       IF #inB15 THEN
           #outR15 := #inR15 * 2.0;
       END_IF;
       // step 536
       #tI36 := #inI16 + #cI26;
       IF #inB16 THEN
           #outR16 := #inR16 * 2.0;
       END_IF;
       // step 537
       #tI37 := #inI17 + #cI27;
       IF #inB17 THEN
           #outR17 := #inR17 * 2.0;
       END_IF;
       // step 538
       #tI38 := #inI18 + #cI28;
       IF #inB18 THEN
           #outR18 := #inR18 * 2.0;
       END_IF;
       // step 539
       #tI39 := #inI19 + #cI29;
       IF #inB19 THEN
           #outR19 := #inR19 * 2.0;
       END_IF;
       // step 540
       #tI40 := #inI20 + #cI0;
       IF #inB20 THEN
           #outR0 := #inR0 * 2.0;
       END_IF;
       // step 541
       #tI41 := #inI21 + #cI1;
       IF #inB21 THEN
           #outR1 := #inR1 * 2.0;
       END_IF;
       // step 542
       #tI42 := #inI22 + #cI2;
       IF #inB22 THEN
           #outR2 := #inR2 * 2.0;
       END_IF;
       // step 543
       #tI43 := #inI23 + #cI3;
       IF #inB23 THEN
           #outR3 := #inR3 * 2.0;
       END_IF;
       // step 544
       #tI44 := #inI24 + #cI4;
       IF #inB24 THEN
           #outR4 := #inR4 * 2.0;
       END_IF;
       // step 545
       #tI45 := #inI25 + #cI5;
       IF #inB25 THEN
           #outR5 := #inR5 * 2.0;
       END_IF;
       // step 546
       #tI46 := #inI26 + #cI6;
       IF #inB26 THEN
           #outR6 := #inR6 * 2.0;
       END_IF;
       // step 547
       #tI47 := #inI27 + #cI7;
       IF #inB27 THEN
           #outR7 := #inR7 * 2.0;
       END_IF;
       // step 548
       #tI48 := #inI28 + #cI8;
       IF #inB28 THEN
           #outR8 := #inR8 * 2.0;
       END_IF;
       // step 549
       #tI49 := #inI29 + #cI9;
       IF #inB29 THEN
           #outR9 := #inR9 * 2.0;
       END_IF;
       END_REGION
       REGION part 11
       // step 550
       #tI50 := #inI30 + #cI10;
       IF #inB30 THEN
           #outR10 := #inR10 * 2.0;
       END_IF;
       // step 551
       #tI51 := #inI31 + #cI11;
       IF #inB31 THEN
           #outR11 := #inR11 * 2.0;
       END_IF;
       // step 552
       #tI52 := #inI32 + #cI12;
       IF #inB32 THEN
           #outR12 := #inR12 * 2.0;
       END_IF;
       // step 553
       #tI53 := #inI33 + #cI13;
       IF #inB33 THEN
           #outR13 := #inR13 * 2.0;
       END_IF;
       // step 554
       #tI54 := #inI34 + #cI14;
       IF #inB34 THEN
           #outR14 := #inR14 * 2.0;
       END_IF;
       // step 555
       #tI55 := #inI35 + #cI15;
       IF #inB35 THEN
           #outR15 := #inR15 * 2.0;
       END_IF;
       // step 556
       #tI56 := #inI36 + #cI16;
       IF #inB36 THEN
           #outR16 := #inR16 * 2.0;
       END_IF;
       // step 557
       #tI57 := #inI37 + #cI17;
       IF #inB37 THEN
           #outR17 := #inR17 * 2.0;
       END_IF;
       // step 558
       #tI58 := #inI38 + #cI18;
       IF #inB38 THEN
           #outR18 := #inR18 * 2.0;
       END_IF;
       // step 559
       #tI59 := #inI39 + #cI19;
       IF #inB39 THEN
           #outR19 := #inR19 * 2.0;
       END_IF;
       // step 560
       #tI60 := #inI0 + #cI20;
       IF #inB0 THEN
           #outR0 := #inR0 * 2.0;
       END_IF;
       // step 561
       #tI61 := #inI1 + #cI21;
       IF #inB1 THEN
           #outR1 := #inR1 * 2.0;
       END_IF;
       // step 562
       #tI62 := #inI2 + #cI22;
       IF #inB2 THEN
           #outR2 := #inR2 * 2.0;
       END_IF;
       // step 563
       #tI63 := #inI3 + #cI23;
       IF #inB3 THEN
           #outR3 := #inR3 * 2.0;
       END_IF;
       // step 564
       #tI64 := #inI4 + #cI24;
       IF #inB4 THEN
           #outR4 := #inR4 * 2.0;
       END_IF;
       // step 565
       #tI65 := #inI5 + #cI25;
       IF #inB5 THEN
           #outR5 := #inR5 * 2.0;
       END_IF;
       // step 566
       #tI66 := #inI6 + #cI26;
       IF #inB6 THEN
           #outR6 := #inR6 * 2.0;
       END_IF;
       // step 567
       #tI67 := #inI7 + #cI27;
       IF #inB7 THEN
           #outR7 := #inR7 * 2.0;
       END_IF;
       // step 568
       #tI68 := #inI8 + #cI28;
       IF #inB8 THEN
           #outR8 := #inR8 * 2.0;
       END_IF;
       // step 569
       #tI69 := #inI9 + #cI29;
       IF #inB9 THEN
           #outR9 := #inR9 * 2.0;
       END_IF;
       // step 570
       #tI70 := #inI10 + #cI0;
       IF #inB10 THEN
           #outR10 := #inR10 * 2.0;
       END_IF;
       // step 571
       #tI71 := #inI11 + #cI1;
       IF #inB11 THEN
           #outR11 := #inR11 * 2.0;
       END_IF;
       // step 572
       #tI72 := #inI12 + #cI2;
       IF #inB12 THEN
           #outR12 := #inR12 * 2.0;
       END_IF;
       // step 573
       #tI73 := #inI13 + #cI3;
       IF #inB13 THEN
           #outR13 := #inR13 * 2.0;
       END_IF;
       // step 574
       #tI74 := #inI14 + #cI4;
       IF #inB14 THEN
           #outR14 := #inR14 * 2.0;
       END_IF;
       // step 575
       #tI75 := #inI15 + #cI5;
       IF #inB15 THEN
           #outR15 := #inR15 * 2.0;
       END_IF;
       // step 576
       #tI76 := #inI16 + #cI6;
       IF #inB16 THEN
           #outR16 := #inR16 * 2.0;
       END_IF;
       // step 577
       #tI77 := #inI17 + #cI7;
       IF #inB17 THEN
           #outR17 := #inR17 * 2.0;
       END_IF;
       // step 578
       #tI78 := #inI18 + #cI8;
       IF #inB18 THEN
           #outR18 := #inR18 * 2.0;
       END_IF;
       // step 579
       #tI79 := #inI19 + #cI9;
       IF #inB19 THEN
           #outR19 := #inR19 * 2.0;
       END_IF;
       // step 580
       #tI80 := #inI20 + #cI10;
       IF #inB20 THEN
           #outR0 := #inR0 * 2.0;
       END_IF;
       // step 581
       #tI81 := #inI21 + #cI11;
       IF #inB21 THEN
           #outR1 := #inR1 * 2.0;
       END_IF;
       // step 582
       #tI82 := #inI22 + #cI12;
       IF #inB22 THEN
           #outR2 := #inR2 * 2.0;
       END_IF;
       // step 583
       #tI83 := #inI23 + #cI13;
       IF #inB23 THEN
           #outR3 := #inR3 * 2.0;
       END_IF;
       // step 584
       #tI84 := #inI24 + #cI14;
       IF #inB24 THEN
           #outR4 := #inR4 * 2.0;
       END_IF;
       // step 585
       #tI85 := #inI25 + #cI15;
       IF #inB25 THEN
           #outR5 := #inR5 * 2.0;
       END_IF;
       // step 586
       #tI86 := #inI26 + #cI16;
       IF #inB26 THEN
           #outR6 := #inR6 * 2.0;
       END_IF;
       // step 587
       #tI87 := #inI27 + #cI17;
       IF #inB27 THEN
           #outR7 := #inR7 * 2.0;
       END_IF;
       // step 588
       #tI88 := #inI28 + #cI18;
       IF #inB28 THEN
           #outR8 := #inR8 * 2.0;
       END_IF;
       // step 589
       #tI89 := #inI29 + #cI19;
       IF #inB29 THEN
           #outR9 := #inR9 * 2.0;
       END_IF;
       // step 590
       #tI90 := #inI30 + #cI20;
       IF #inB30 THEN
           #outR10 := #inR10 * 2.0;
       END_IF;
       // step 591
       #tI91 := #inI31 + #cI21;
       IF #inB31 THEN
           #outR11 := #inR11 * 2.0;
       END_IF;
       // step 592
       #tI92 := #inI32 + #cI22;
       IF #inB32 THEN
           #outR12 := #inR12 * 2.0;
       END_IF;
       // step 593
       #tI93 := #inI33 + #cI23;
       IF #inB33 THEN
           #outR13 := #inR13 * 2.0;
       END_IF;
       // step 594
       #tI94 := #inI34 + #cI24;
       IF #inB34 THEN
           #outR14 := #inR14 * 2.0;
       END_IF;
       // step 595
       #tI95 := #inI35 + #cI25;
       IF #inB35 THEN
           #outR15 := #inR15 * 2.0;
       END_IF;
       // step 596
       #tI96 := #inI36 + #cI26;
       IF #inB36 THEN
           #outR16 := #inR16 * 2.0;
       END_IF;
       // step 597
       #tI97 := #inI37 + #cI27;
       IF #inB37 THEN
           #outR17 := #inR17 * 2.0;
       END_IF;
       // step 598
       #tI98 := #inI38 + #cI28;
       IF #inB38 THEN
           #outR18 := #inR18 * 2.0;
       END_IF;
       // step 599
       #tI99 := #inI39 + #cI29;
       IF #inB39 THEN
           #outR19 := #inR19 * 2.0;
       END_IF;
       END_REGION
END_FUNCTION_BLOCK

FUNCTION_BLOCK "FB_MixedStl"   // FB900, LAD
{ S7_Optimized_Access := 'TRUE' }
VERSION : 0.1
   VAR_INPUT
      inB0 : Bool;   // input bit 0
      inB1 : Bool;
      inB2 : Bool;
      inB3 : Bool;
      inB4 : Bool;
      inB5 : Bool;
      inB6 : Bool;
      inB7 : Bool;
      inB8 : Bool;
      inB9 : Bool;
      inB10 : Bool;   // input bit 10
      inB11 : Bool;
      inB12 : Bool;
      inB13 : Bool;
      inB14 : Bool;
      inB15 : Bool;
      inB16 : Bool;
      inB17 : Bool;
      inB18 : Bool;
      inB19 : Bool;
      inB20 : Bool;   // input bit 20
      inB21 : Bool;
      inB22 : Bool;
      inB23 : Bool;
      inB24 : Bool;
      inB25 : Bool;
      inB26 : Bool;
      inB27 : Bool;
      inB28 : Bool;
      inB29 : Bool;
      inB30 : Bool;   // input bit 30
      inB31 : Bool;
      inB32 : Bool;
      inB33 : Bool;
      inB34 : Bool;
      inB35 : Bool;
      inB36 : Bool;
      inB37 : Bool;
      inB38 : Bool;
      inB39 : Bool;
      inI0 : Int;
      inI1 : Int;
      inI2 : Int;
      inI3 : Int;
      inI4 : Int;
      inI5 : Int;
      inI6 : Int;
      inI7 : Int;
      inI8 : Int;
      inI9 : Int;
      inI10 : Int;
      inI11 : Int;
      inI12 : Int;
      inI13 : Int;
      inI14 : Int;
      inI15 : Int;
      inI16 : Int;
      inI17 : Int;
      inI18 : Int;
      inI19 : Int;
      inI20 : Int;
      inI21 : Int;
      inI22 : Int;
      inI23 : Int;
      inI24 : Int;
      inI25 : Int;
      inI26 : Int;
      inI27 : Int;
      inI28 : Int;
      inI29 : Int;
      inI30 : Int;
      inI31 : Int;
      inI32 : Int;
      inI33 : Int;
      inI34 : Int;
      inI35 : Int;
      inI36 : Int;
      inI37 : Int;
      inI38 : Int;
      inI39 : Int;
      inR0 : Real;
      inR1 : Real;
      inR2 : Real;
      inR3 : Real;
      inR4 : Real;
      inR5 : Real;
      inR6 : Real;
      inR7 : Real;
      inR8 : Real;
      inR9 : Real;
      inR10 : Real;
      inR11 : Real;
      inR12 : Real;
      inR13 : Real;
      inR14 : Real;
      inR15 : Real;
      inR16 : Real;
      inR17 : Real;
      inR18 : Real;
      inR19 : Real;
      inD0 : DInt;
      inD1 : DInt;
      inD2 : DInt;
      inD3 : DInt;
      inD4 : DInt;
      inD5 : DInt;
      inD6 : DInt;
      inD7 : DInt;
      inD8 : DInt;
      inD9 : DInt;
      inD10 : DInt;
      inD11 : DInt;
      inD12 : DInt;
      inD13 : DInt;
      inD14 : DInt;
      inD15 : DInt;
      inD16 : DInt;
      inD17 : DInt;
      inD18 : DInt;
      inD19 : DInt;
      inArr : Array[0..99] of Int;   // input array
      inStr : String[40];
      inSt : Struct
         x : Int;
         y : Real;
         z : Bool;
      END_STRUCT;
   END_VAR
   VAR_OUTPUT
      outB0 : Bool;
      outB1 : Bool;
      outB2 : Bool;
      outB3 : Bool;
      outB4 : Bool;
      outB5 : Bool;
      outB6 : Bool;
      outB7 : Bool;
      outB8 : Bool;
      outB9 : Bool;
      outB10 : Bool;
      outB11 : Bool;
      outB12 : Bool;
      outB13 : Bool;
      outB14 : Bool;
      outB15 : Bool;
      outB16 : Bool;
      outB17 : Bool;
      outB18 : Bool;
      outB19 : Bool;
      outB20 : Bool;
      outB21 : Bool;
      outB22 : Bool;
      outB23 : Bool;
      outB24 : Bool;
      outB25 : Bool;
      outB26 : Bool;
      outB27 : Bool;
      outB28 : Bool;
      outB29 : Bool;
      outB30 : Bool;
      outB31 : Bool;
      outB32 : Bool;
      outB33 : Bool;
      outB34 : Bool;
      outB35 : Bool;
      outB36 : Bool;
      outB37 : Bool;
      outB38 : Bool;
      outB39 : Bool;
      outI0 : Int;   // output int 0
      outI1 : Int;
      outI2 : Int;
      outI3 : Int;
      outI4 : Int;
      outI5 : Int;
      outI6 : Int;
      outI7 : Int;
      outI8 : Int;
      outI9 : Int;
      outI10 : Int;   // output int 10
      outI11 : Int;
      outI12 : Int;
      outI13 : Int;
      outI14 : Int;
      outI15 : Int;
      outI16 : Int;
      outI17 : Int;
      outI18 : Int;
      outI19 : Int;
      outI20 : Int;   // output int 20
      outI21 : Int;
      outI22 : Int;
      outI23 : Int;
      outI24 : Int;
      outI25 : Int;
      outI26 : Int;
      outI27 : Int;
      outI28 : Int;
      outI29 : Int;
      outI30 : Int;   // output int 30
      outI31 : Int;
      outI32 : Int;
      outI33 : Int;
      outI34 : Int;
      outI35 : Int;
      outI36 : Int;
      outI37 : Int;
      outI38 : Int;
      outI39 : Int;
      outR0 : Real;
      outR1 : Real;
      outR2 : Real;
      outR3 : Real;
      outR4 : Real;
      outR5 : Real;
      outR6 : Real;
      outR7 : Real;
      outR8 : Real;
      outR9 : Real;
      outR10 : Real;
      outR11 : Real;
      outR12 : Real;
      outR13 : Real;
      outR14 : Real;
      outR15 : Real;
      outR16 : Real;
      outR17 : Real;
      outR18 : Real;
      outR19 : Real;
      outD0 : DInt;
      outD1 : DInt;
      outD2 : DInt;
      outD3 : DInt;
      outD4 : DInt;
      outD5 : DInt;
      outD6 : DInt;
      outD7 : DInt;
      outD8 : DInt;
      outD9 : DInt;
      outD10 : DInt;
      outD11 : DInt;
      outD12 : DInt;
      outD13 : DInt;
      outD14 : DInt;
      outD15 : DInt;
      outD16 : DInt;
      outD17 : DInt;
      outD18 : DInt;
      outD19 : DInt;
   END_VAR
   VAR_IN_OUT
      ioI0 : Int;
      ioI1 : Int;
      ioI2 : Int;
      ioI3 : Int;
      ioI4 : Int;
      ioI5 : Int;
      ioI6 : Int;
      ioI7 : Int;
      ioI8 : Int;
      ioI9 : Int;
      ioI10 : Int;
      ioI11 : Int;
      ioI12 : Int;
      ioI13 : Int;
      ioI14 : Int;
      ioI15 : Int;
      ioI16 : Int;
      ioI17 : Int;
      ioI18 : Int;
      ioI19 : Int;
      ioI20 : Int;
      ioI21 : Int;
      ioI22 : Int;
      ioI23 : Int;
      ioI24 : Int;
      ioI25 : Int;
      ioI26 : Int;
      ioI27 : Int;
      ioI28 : Int;
      ioI29 : Int;
      ioI30 : Int;
      ioI31 : Int;
      ioI32 : Int;
      ioI33 : Int;
      ioI34 : Int;
      ioI35 : Int;
      ioI36 : Int;
      ioI37 : Int;
      ioI38 : Int;
      ioI39 : Int;
      ioI40 : Int;
      ioI41 : Int;
      ioI42 : Int;
      ioI43 : Int;
      ioI44 : Int;
      ioI45 : Int;
      ioI46 : Int;
      ioI47 : Int;
      ioI48 : Int;
      ioI49 : Int;
      ioI50 : Int;
      ioI51 : Int;
      ioI52 : Int;
      ioI53 : Int;
      ioI54 : Int;
      ioI55 : Int;
      ioI56 : Int;
      ioI57 : Int;
      ioI58 : Int;
      ioI59 : Int;
   END_VAR
   VAR
      stI0 : Int := 0;   // static 0
      stI1 : Int;
      stI2 : Int;
      stI3 : Int;
      stI4 : Int;
      stI5 : Int;
      stI6 : Int;
      stI7 : Int := 7;
      stI8 : Int;
      stI9 : Int;
      stI10 : Int;
      stI11 : Int;
      stI12 : Int;
      stI13 : Int;
      stI14 : Int := 14;
      stI15 : Int;
      stI16 : Int;
      stI17 : Int;
      stI18 : Int;
      stI19 : Int;
      stI20 : Int;
      stI21 : Int := 21;
      stI22 : Int;
      stI23 : Int;
      stI24 : Int;
      stI25 : Int;   // static 25
      stI26 : Int;
      stI27 : Int;
      stI28 : Int := 28;
      stI29 : Int;
      stI30 : Int;
      stI31 : Int;
      stI32 : Int;
      stI33 : Int;
      stI34 : Int;
      stI35 : Int := 35;
      stI36 : Int;
      stI37 : Int;
      stI38 : Int;
      stI39 : Int;
      stI40 : Int;
      stI41 : Int;
      stI42 : Int := 42;
      stI43 : Int;
      stI44 : Int;
      stI45 : Int;
      stI46 : Int;
      stI47 : Int;
      stI48 : Int;
      stI49 : Int := 49;
      stI50 : Int;   // static 50
      stI51 : Int;
      stI52 : Int;
      stI53 : Int;
      stI54 : Int;
      stI55 : Int;
      stI56 : Int := 56;
      stI57 : Int;
      stI58 : Int;
      stI59 : Int;
      stI60 : Int;
      stI61 : Int;
      stI62 : Int;
      stI63 : Int := 63;
      stI64 : Int;
      stI65 : Int;
      stI66 : Int;
      stI67 : Int;
      stI68 : Int;
      stI69 : Int;
      stI70 : Int := 70;
      stI71 : Int;
      stI72 : Int;
      stI73 : Int;
      stI74 : Int;
      stI75 : Int;   // static 75
      stI76 : Int;
      stI77 : Int := 77;
      stI78 : Int;
      stI79 : Int;
      stI80 : Int;
      stI81 : Int;
      stI82 : Int;
      stI83 : Int;
      stI84 : Int := 84;
      stI85 : Int;
      stI86 : Int;
      stI87 : Int;
      stI88 : Int;
      stI89 : Int;
      stI90 : Int;
      stI91 : Int := 91;
      stI92 : Int;
      stI93 : Int;
      stI94 : Int;
      stI95 : Int;
      stI96 : Int;
      stI97 : Int;
      stI98 : Int := 98;
      stI99 : Int;
      stI100 : Int;   // static 100
      stI101 : Int;
      stI102 : Int;
      stI103 : Int;
      stI104 : Int;
      stI105 : Int := 105;
      stI106 : Int;
      stI107 : Int;
      stI108 : Int;
      stI109 : Int;
      stI110 : Int;
      stI111 : Int;
      stI112 : Int := 112;
      stI113 : Int;
      stI114 : Int;
      stI115 : Int;
      stI116 : Int;
      stI117 : Int;
      stI118 : Int;
      stI119 : Int := 119;
      stI120 : Int;
      stI121 : Int;
      stI122 : Int;
      stI123 : Int;
      stI124 : Int;
      stI125 : Int;   // static 125
      stI126 : Int := 126;
      stI127 : Int;
      stI128 : Int;
      stI129 : Int;
      stI130 : Int;
      stI131 : Int;
      stI132 : Int;
      stI133 : Int := 133;
      stI134 : Int;
      stI135 : Int;
      stI136 : Int;
      stI137 : Int;
      stI138 : Int;
      stI139 : Int;
      stI140 : Int := 140;
      stI141 : Int;
      stI142 : Int;
      stI143 : Int;
      stI144 : Int;
      stI145 : Int;
      stI146 : Int;
      stI147 : Int := 147;
      stI148 : Int;
      stI149 : Int;
      stI150 : Int;   // static 150
      stI151 : Int;
      stI152 : Int;
      stI153 : Int;
      stI154 : Int := 154;
      stI155 : Int;
      stI156 : Int;
      stI157 : Int;
      stI158 : Int;
      stI159 : Int;
      stI160 : Int;
      stI161 : Int := 161;
      stI162 : Int;
      stI163 : Int;
      stI164 : Int;
      stI165 : Int;
      stI166 : Int;
      stI167 : Int;
      stI168 : Int := 168;
      stI169 : Int;
      stI170 : Int;
      stI171 : Int;
      stI172 : Int;
      stI173 : Int;
      stI174 : Int;
      stI175 : Int := 175;   // static 175
      stI176 : Int;
      stI177 : Int;
      stI178 : Int;
      stI179 : Int;
      stI180 : Int;
      stI181 : Int;
      stI182 : Int := 182;
      stI183 : Int;
      stI184 : Int;
      stI185 : Int;
      stI186 : Int;
      stI187 : Int;
      stI188 : Int;
      stI189 : Int := 189;
      stI190 : Int;
      stI191 : Int;
      stI192 : Int;
      stI193 : Int;
      stI194 : Int;
      stI195 : Int;
      stI196 : Int := 196;
      stI197 : Int;
      stI198 : Int;
      stI199 : Int;
      stB0 : Bool := TRUE;
      stB1 : Bool;
      stB2 : Bool;
      stB3 : Bool := TRUE;
      stB4 : Bool;
      stB5 : Bool;
      stB6 : Bool := TRUE;
      stB7 : Bool;
      stB8 : Bool;
      stB9 : Bool := TRUE;
      stB10 : Bool;
      stB11 : Bool;
      stB12 : Bool := TRUE;
      stB13 : Bool;
      stB14 : Bool;
      stB15 : Bool := TRUE;
      stB16 : Bool;
      stB17 : Bool;
      stB18 : Bool := TRUE;
      stB19 : Bool;
      stB20 : Bool;
      stB21 : Bool := TRUE;
      stB22 : Bool;
      stB23 : Bool;
      stB24 : Bool := TRUE;
      stB25 : Bool;
      stB26 : Bool;
      stB27 : Bool := TRUE;
      stB28 : Bool;
      stB29 : Bool;
      stB30 : Bool := TRUE;
      stB31 : Bool;
      stB32 : Bool;
      stB33 : Bool := TRUE;
      stB34 : Bool;
      stB35 : Bool;
      stB36 : Bool := TRUE;
      stB37 : Bool;
      stB38 : Bool;
      stB39 : Bool := TRUE;
      stB40 : Bool;
      stB41 : Bool;
      stB42 : Bool := TRUE;
      stB43 : Bool;
      stB44 : Bool;
      stB45 : Bool := TRUE;
      stB46 : Bool;
      stB47 : Bool;
      stB48 : Bool := TRUE;
      stB49 : Bool;
      stB50 : Bool;
      stB51 : Bool := TRUE;
      stB52 : Bool;
      stB53 : Bool;
      stB54 : Bool := TRUE;
      stB55 : Bool;
      stB56 : Bool;
      stB57 : Bool := TRUE;
      stB58 : Bool;
      stB59 : Bool;
      stB60 : Bool := TRUE;
      stB61 : Bool;
      stB62 : Bool;
      stB63 : Bool := TRUE;
      stB64 : Bool;
      stB65 : Bool;
      stB66 : Bool := TRUE;
      stB67 : Bool;
      stB68 : Bool;
      stB69 : Bool := TRUE;
      stB70 : Bool;
      stB71 : Bool;
      stB72 : Bool := TRUE;
      stB73 : Bool;
      stB74 : Bool;
      stB75 : Bool := TRUE;
      stB76 : Bool;
      stB77 : Bool;
      stB78 : Bool := TRUE;
      stB79 : Bool;
      stB80 : Bool;
      stB81 : Bool := TRUE;
      stB82 : Bool;
      stB83 : Bool;
      stB84 : Bool := TRUE;
      stB85 : Bool;
      stB86 : Bool;
      stB87 : Bool := TRUE;
      stB88 : Bool;
      stB89 : Bool;
      stB90 : Bool := TRUE;
      stB91 : Bool;
      stB92 : Bool;
      stB93 : Bool := TRUE;
      stB94 : Bool;
      stB95 : Bool;
      stB96 : Bool := TRUE;
      stB97 : Bool;
      stB98 : Bool;
      stB99 : Bool := TRUE;
      stArr : Array[1..10, 0..4] of Real;
      stSt : Struct
         "a" : Int;
         "b" : Array[0..3] of Bool;
         c : Time;
      END_STRUCT;
   END_VAR
   VAR_TEMP
      tI0 : Int;
      tI1 : Int;
      tI2 : Int;
      tI3 : Int;
      tI4 : Int;
      tI5 : Int;
      tI6 : Int;
      tI7 : Int;
      tI8 : Int;
      tI9 : Int;
      tI10 : Int;
      tI11 : Int;
      tI12 : Int;
      tI13 : Int;
      tI14 : Int;
      tI15 : Int;
      tI16 : Int;
      tI17 : Int;
      tI18 : Int;
      tI19 : Int;
      tI20 : Int;
      tI21 : Int;
      tI22 : Int;
      tI23 : Int;
      tI24 : Int;
      tI25 : Int;
      tI26 : Int;
      tI27 : Int;
      tI28 : Int;
      tI29 : Int;
      tI30 : Int;
      tI31 : Int;
      tI32 : Int;
      tI33 : Int;
      tI34 : Int;
      tI35 : Int;
      tI36 : Int;
      tI37 : Int;
      tI38 : Int;
      tI39 : Int;
      tI40 : Int;
      tI41 : Int;
      tI42 : Int;
      tI43 : Int;
      tI44 : Int;
      tI45 : Int;
      tI46 : Int;
      tI47 : Int;
      tI48 : Int;
      tI49 : Int;
      tI50 : Int;
      tI51 : Int;
      tI52 : Int;
      tI53 : Int;
      tI54 : Int;
      tI55 : Int;
      tI56 : Int;
      tI57 : Int;
      tI58 : Int;
      tI59 : Int;
      tI60 : Int;
      tI61 : Int;
      tI62 : Int;
      tI63 : Int;
      tI64 : Int;
      tI65 : Int;
      tI66 : Int;
      tI67 : Int;
      tI68 : Int;
      tI69 : Int;
      tI70 : Int;
      tI71 : Int;
      tI72 : Int;
      tI73 : Int;
      tI74 : Int;
      tI75 : Int;
      tI76 : Int;
      tI77 : Int;
      tI78 : Int;
      tI79 : Int;
      tI80 : Int;
      tI81 : Int;
      tI82 : Int;
      tI83 : Int;
      tI84 : Int;
      tI85 : Int;
      tI86 : Int;
      tI87 : Int;
      tI88 : Int;
      tI89 : Int;
      tI90 : Int;
      tI91 : Int;
      tI92 : Int;
      tI93 : Int;
      tI94 : Int;
      tI95 : Int;
      tI96 : Int;
      tI97 : Int;
      tI98 : Int;
      tI99 : Int;
      tR0 : Real;
      tR1 : Real;
      tR2 : Real;
      tR3 : Real;
      tR4 : Real;
      tR5 : Real;
      tR6 : Real;
      tR7 : Real;
      tR8 : Real;
      tR9 : Real;
      tR10 : Real;
      tR11 : Real;
      tR12 : Real;
      tR13 : Real;
      tR14 : Real;
      tR15 : Real;
      tR16 : Real;
      tR17 : Real;
      tR18 : Real;
      tR19 : Real;
      tR20 : Real;
      tR21 : Real;
      tR22 : Real;
      tR23 : Real;
      tR24 : Real;
      tR25 : Real;
      tR26 : Real;
      tR27 : Real;
      tR28 : Real;
      tR29 : Real;
      tR30 : Real;
      tR31 : Real;
      tR32 : Real;
      tR33 : Real;
      tR34 : Real;
      tR35 : Real;
      tR36 : Real;
      tR37 : Real;
      tR38 : Real;
      tR39 : Real;
      tR40 : Real;
      tR41 : Real;
      tR42 : Real;
      tR43 : Real;
      tR44 : Real;
      tR45 : Real;
      tR46 : Real;
      tR47 : Real;
      tR48 : Real;
      tR49 : Real;
   END_VAR
   VAR CONSTANT
      cI0 : Int := 0;
      cI1 : Int := 3;
      cI2 : Int := 6;
      cI3 : Int := 9;
      cI4 : Int := 12;
      cI5 : Int := 15;
      cI6 : Int := 18;
      cI7 : Int := 21;
      cI8 : Int := 24;
      cI9 : Int := 27;
      cI10 : Int := 30;
      cI11 : Int := 33;
      cI12 : Int := 36;
      cI13 : Int := 39;
      cI14 : Int := 42;
      cI15 : Int := 45;
      cI16 : Int := 48;
      cI17 : Int := 51;
      cI18 : Int := 54;
      cI19 : Int := 57;
      cI20 : Int := 60;
      cI21 : Int := 63;
      cI22 : Int := 66;
      cI23 : Int := 69;
      cI24 : Int := 72;
      cI25 : Int := 75;
      cI26 : Int := 78;
      cI27 : Int := 81;
      cI28 : Int := 84;
      cI29 : Int := 87;
   END_VAR
BEGIN

REGION Network 1: LAD network 1
   // mixed 1
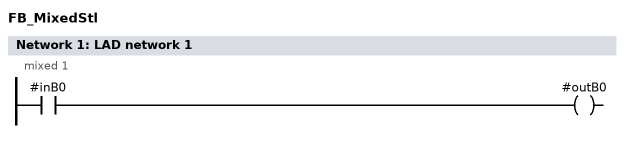
   RUNG wire#powerrail
      Contact( #inB0 )
      Coil( #outB0 )
   END_RUNG
   // the same network as SCL:
   #outB0 := #inB0;
END_REGION

REGION Network 2 (FBD): FBD network 2
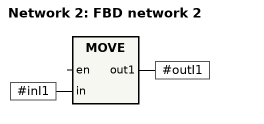
   #outI1 := #inI1;
END_REGION

REGION Network 3 (SCL): SCL network 3
   #tI2 := #inI2 + #cI2;
           IF #inB2 THEN
               #outR2 := #inR2 * 2.0;
           END_IF;
END_REGION

REGION Network 4 (STL): STL network 1
   // comment of STL network 1
         A     #inB0;
         AN    #stB0;
         =     #outB0;
END_REGION

REGION Network 5: LAD network 4
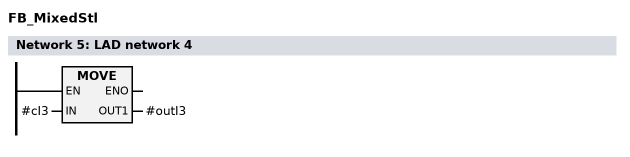
   RUNG wire#powerrail
      Move(in := #cI3, out1 => #outI3)
   END_RUNG
   // the same network as SCL:
   #outI3 := #cI3;
END_REGION

REGION Network 6 (FBD): FBD network 5
   // mixed 5
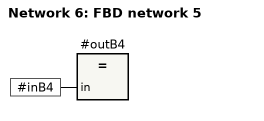
   #outB4 := #inB4;
END_REGION

REGION Network 7 (SCL): SCL network 6
   #tI5 := #inI5 + #cI5;
           IF #inB5 THEN
               #outR5 := #inR5 * 2.0;
           END_IF;
END_REGION

REGION Network 8 (STL): STL network 2
         L     #inI1;
         L     #stI1;
         +I;
         T     #outI1;
END_REGION

REGION Network 9: LAD network 7
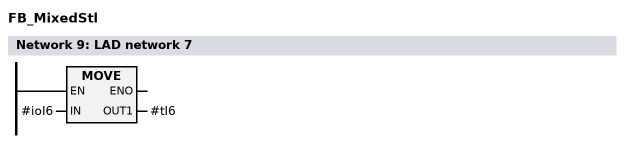
   RUNG wire#powerrail
      Move(in := #ioI6, out1 => #tI6)
   END_RUNG
   // the same network as SCL:
   #tI6 := #ioI6;
END_REGION

REGION Network 10 (FBD): FBD network 8
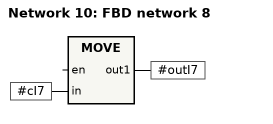
   #outI7 := #cI7;
END_REGION

REGION Network 11 (SCL): SCL network 9
   // mixed 9
   #tI8 := #inI8 + #cI8;
           IF #inB8 THEN
               #outR8 := #inR8 * 2.0;
           END_IF;
END_REGION

REGION Network 12 (STL): STL network 3
         L     #inR2;
         L     #tR2;
         *R;
         T     #outR2;  // product
END_REGION

REGION Network 13: LAD network 10
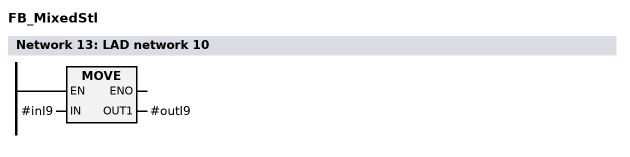
   RUNG wire#powerrail
      Move(in := #inI9, out1 => #outI9)
   END_RUNG
   // the same network as SCL:
   #outI9 := #inI9;
END_REGION

REGION Network 14 (FBD): FBD network 11
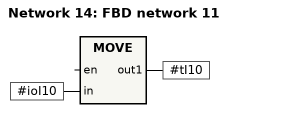
   #tI10 := #ioI10;
END_REGION

REGION Network 15 (SCL): SCL network 12
   #tI11 := #inI11 + #cI11;
           IF #inB11 THEN
               #outR11 := #inR11 * 2.0;
           END_IF;
END_REGION

REGION Network 16 (STL): STL network 4
         A     #inB3;
         AN    #stB3;
         =     #outB3;
END_REGION

REGION Network 17: LAD network 13
   // mixed 13
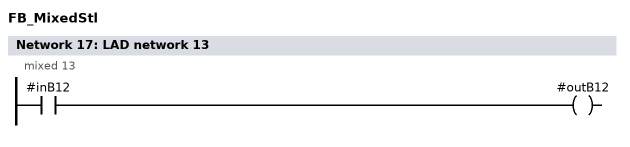
   RUNG wire#powerrail
      Contact( #inB12 )
      Coil( #outB12 )
   END_RUNG
   // the same network as SCL:
   #outB12 := #inB12;
END_REGION

REGION Network 18 (FBD): FBD network 14
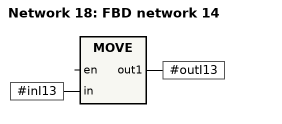
   #outI13 := #inI13;
END_REGION

REGION Network 19 (SCL): SCL network 15
   #tI14 := #inI14 + #cI14;
           IF #inB14 THEN
               #outR14 := #inR14 * 2.0;
           END_IF;
END_REGION

REGION Network 20 (STL): STL network 5
         L     #inI4;
         L     #stI4;
         +I;
         T     #outI4;
END_REGION

REGION Network 21: LAD network 16
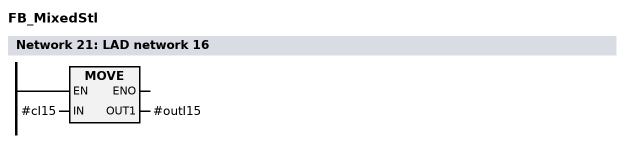
   RUNG wire#powerrail
      Move(in := #cI15, out1 => #outI15)
   END_RUNG
   // the same network as SCL:
   #outI15 := #cI15;
END_REGION

REGION Network 22 (FBD): FBD network 17
   // mixed 17
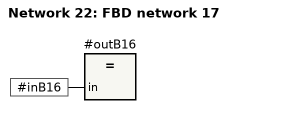
   #outB16 := #inB16;
END_REGION

REGION Network 23 (SCL): SCL network 18
   #tI17 := #inI17 + #cI17;
           IF #inB17 THEN
               #outR17 := #inR17 * 2.0;
           END_IF;
END_REGION

REGION Network 24 (STL): STL network 6
         L     #inR5;
         L     #tR5;
         *R;
         T     #outR5;  // product
END_REGION

REGION Network 25: LAD network 19
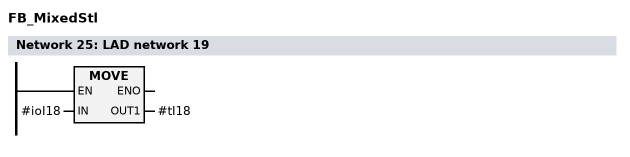
   RUNG wire#powerrail
      Move(in := #ioI18, out1 => #tI18)
   END_RUNG
   // the same network as SCL:
   #tI18 := #ioI18;
END_REGION

REGION Network 26 (FBD): FBD network 20
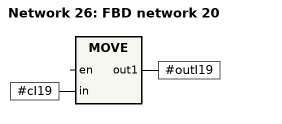
   #outI19 := #cI19;
END_REGION

REGION Network 27 (SCL): SCL network 21
   // mixed 21
   #tI20 := #inI20 + #cI20;
           IF #inB20 THEN
               #outR0 := #inR0 * 2.0;
           END_IF;
END_REGION

REGION Network 28 (STL): STL network 7
         A     #inB6;
         AN    #stB6;
         =     #outB6;
END_REGION

REGION Network 29: LAD network 22
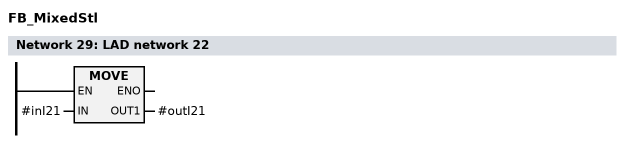
   RUNG wire#powerrail
      Move(in := #inI21, out1 => #outI21)
   END_RUNG
   // the same network as SCL:
   #outI21 := #inI21;
END_REGION

REGION Network 30 (FBD): FBD network 23
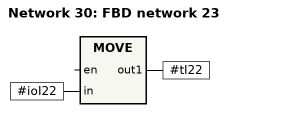
   #tI22 := #ioI22;
END_REGION

REGION Network 31 (SCL): SCL network 24
   #tI23 := #inI23 + #cI23;
           IF #inB23 THEN
               #outR3 := #inR3 * 2.0;
           END_IF;
END_REGION

REGION Network 32 (STL): STL network 8
         L     #inI7;
         L     #stI7;
         +I;
         T     #outI7;
END_REGION

REGION Network 33: LAD network 25
   // mixed 25
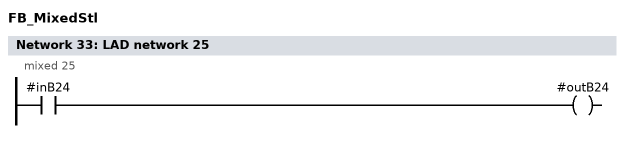
   RUNG wire#powerrail
      Contact( #inB24 )
      Coil( #outB24 )
   END_RUNG
   // the same network as SCL:
   #outB24 := #inB24;
END_REGION

REGION Network 34 (FBD): FBD network 26
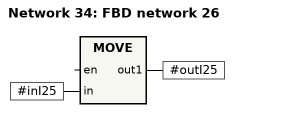
   #outI25 := #inI25;
END_REGION

REGION Network 35 (SCL): SCL network 27
   #tI26 := #inI26 + #cI26;
           IF #inB26 THEN
               #outR6 := #inR6 * 2.0;
           END_IF;
END_REGION

REGION Network 36 (STL): STL network 9
         L     #inR8;
         L     #tR8;
         *R;
         T     #outR8;  // product
END_REGION

REGION Network 37: LAD network 28
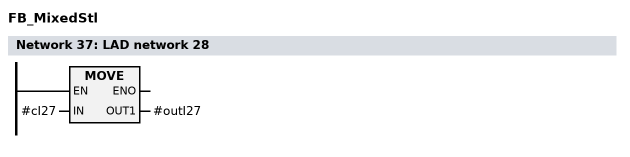
   RUNG wire#powerrail
      Move(in := #cI27, out1 => #outI27)
   END_RUNG
   // the same network as SCL:
   #outI27 := #cI27;
END_REGION

REGION Network 38 (FBD): FBD network 29
   // mixed 29
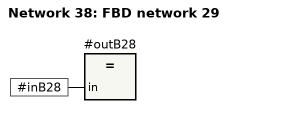
   #outB28 := #inB28;
END_REGION

REGION Network 39 (SCL): SCL network 30
   #tI29 := #inI29 + #cI29;
           IF #inB29 THEN
               #outR9 := #inR9 * 2.0;
           END_IF;
END_REGION

REGION Network 40 (STL): STL network 10
         A     #inB9;
         AN    #stB9;
         =     #outB9;
END_REGION

REGION Network 41: LAD network 31
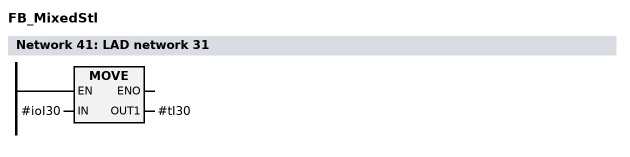
   RUNG wire#powerrail
      Move(in := #ioI30, out1 => #tI30)
   END_RUNG
   // the same network as SCL:
   #tI30 := #ioI30;
END_REGION

REGION Network 42 (FBD): FBD network 32
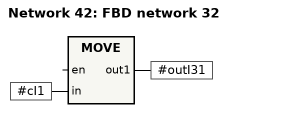
   #outI31 := #cI1;
END_REGION

REGION Network 43 (SCL): SCL network 33
   // mixed 33
   #tI32 := #inI32 + #cI2;
           IF #inB32 THEN
               #outR12 := #inR12 * 2.0;
           END_IF;
END_REGION

REGION Network 44 (STL): STL network 11
   // comment of STL network 11
         L     #inI10;
         L     #stI10;
         +I;
         T     #outI10;
END_REGION

REGION Network 45: LAD network 34
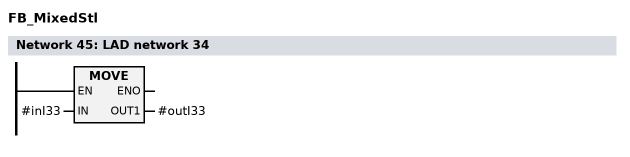
   RUNG wire#powerrail
      Move(in := #inI33, out1 => #outI33)
   END_RUNG
   // the same network as SCL:
   #outI33 := #inI33;
END_REGION

REGION Network 46 (FBD): FBD network 35
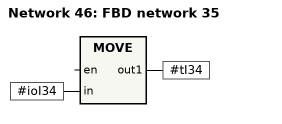
   #tI34 := #ioI34;
END_REGION

REGION Network 47 (SCL): SCL network 36
   #tI35 := #inI35 + #cI5;
           IF #inB35 THEN
               #outR15 := #inR15 * 2.0;
           END_IF;
END_REGION

REGION Network 48 (STL): STL network 12
         L     #inR11;
         L     #tR11;
         *R;
         T     #outR11;  // product
END_REGION

REGION Network 49: LAD network 37
   // mixed 37
